(* IEC 61131-3 sources: kns-pump-station/tests/POUs/Log/FB_TestAlarmSource, 6 files *)

(* ---- FB_TestAlarmSource.decl.st ---- *)
// Назначение: тестовый источник тревог (PL.I_AlarmSource) для FB_AlarmSummary_Test — до восьми PL.FB_Alarm с
//             условиями, номерами и настройками от теста; вызов тела выполняет запросы Ack/Shelve/Unshelve.
// Автор:      kr0nsch
// Версия:     0.1.0
// Документ:   docs/DESIGN.md, разделы 9.3, 14.1
FUNCTION_BLOCK FB_TestAlarmSource IMPLEMENTS PL.I_AlarmSource
VAR_INPUT
    uiSlots   : UINT;               // используемых слотов (AlarmCount), не больше ALM_SLOT_MAX + 1
    udiIdBase : UDINT;              // номер тревоги слота 0
    axIn      : ARRAY[0..GVL_Const.ALM_SLOT_MAX] OF BOOL;              // условия тревог
    astCfg    : ARRAY[0..GVL_Const.ALM_SLOT_MAX] OF PL.ST_AlarmCfg;    // настройки (умолчание — Medium, 8 ч)
    itfTime   : PL.I_TimeSource;    // подменное время теста
END_VAR
VAR
    afbAlarm : ARRAY[0..GVL_Const.ALM_SLOT_MAX] OF PL.FB_Alarm;   // тревоги слотов
    uiK      : UINT;                // номер слота, с 1
END_VAR

(* ---- AckAll.method.decl.st ---- *)
// Квитировать все слоты; TRUE — было что квитировать
METHOD AckAll : BOOL
VAR
    uiI : UINT;                     // номер слота, с 1
END_VAR

(* ---- AckAll.method.impl.st ---- *)
AckAll := FALSE;
FOR uiI := 1 TO MIN(uiSlots, GVL_Const.ALM_SLOT_MAX + 1) DO
    AckAll := afbAlarm[uiI - 1].Ack() OR AckAll;
END_FOR

(* ---- FB_TestAlarmSource.impl.st ---- *)
FOR uiK := 1 TO MIN(uiSlots, GVL_Const.ALM_SLOT_MAX + 1) DO
    afbAlarm[uiK - 1](xIn := axIn[uiK - 1], udiId := udiIdBase + uiK - 1, stCfg := astCfg[uiK - 1], itfTime := itfTime);
END_FOR

(* ---- GetAlarm.method.decl.st ---- *)
// Тревога слота uiIndex; вне 0…AlarmCount - 1 — 0
METHOD GetAlarm : PL.I_Alarm
VAR_INPUT
    uiIndex : UINT;                 // номер слота
END_VAR

(* ---- GetAlarm.method.impl.st ---- *)
IF uiIndex < MIN(uiSlots, GVL_Const.ALM_SLOT_MAX + 1) THEN
    GetAlarm := afbAlarm[uiIndex];
ELSE
    GetAlarm := 0;
END_IF
